Fanuc KAREL source: KA00043.KL

PROGRAM KA00043
%NOLOCKGROUP
VAR
  SRC: STRING[80]
  DST: XYZWPREXT
BEGIN
  SRC = 'A'
  DST = SRC
END KA00043
